(* IEC 61131-3 sources: T4Exjobb/Sigma/Stations/MachineControl/MachineControl/Network, 1 file *)

(* ---- ConfigObjects.st ---- *)
FUNCTION GLOBAL TAB TASK_CONF
_K_TASK, _K_REAL,
_K_END_VAR,

_K_TASK, _K_CYCLIC,
_K_END_VAR,

_K_TASK, _K_BACKGROUND,
_K_END_VAR,

_K_END_CONF
END_FUNCTION

FUNCTION GLOBAL TAB IPR_CONF
_K_IPR
	0$UINT,
_K_END_VAR,
_K_END_CONF
END_FUNCTION

FUNCTION GLOBAL TAB CONFIG_TABLES
00034$UINT,
0$UINT, 0, 11, "_ALARMX0PARA",
0$UINT, 0, 19, "_ALARMXBUFFER",
0$UINT, 1, 3, "_CHECKONLINESTATUS",
0$UINT, 1, 0, "_CHECKSUM",
0$UINT, 1, 1, "_MULTITASK",
0$UINT, 1, 0, "_SIG_LSL_CMULTIMASTERSTATE",
0$UINT, 0, 0, "_STDLIB",
0$UINT, 2, 0, "_SYNCTIMEPLC",
0$UINT, 0, 7, "_SYSDATETIME",
0$UINT, 0, 0, "_SYSDATETIME2",
0$UINT, 1, 1, "_TASKOBJECTCONTROL",
0$UINT, 1, 17, "_TCPIP_CLIENT",
0$UINT, 1, 36, "_TCPIP_SERVER",
0$UINT, 1, 20, "ASCII_BIN",
0$UINT, 0, 4, "CRITICALSECTION",
0$UINT, 1, 0, "DATAMANAGER",
0$UINT, 1, 0, "DATAMANAGERFIFO",
0$UINT, 1, 0, "DATAMANAGERPRIORITY",
0$UINT, 1, 2, "GETOSVERSION",
0$UINT, 0, 2, "GETTASKHANDLE",
0$UINT, 1, 22, "MERKEREX",
0$UINT, 1, 68, "PLC_INFO",
0$UINT, 1, 3, "RAM",
0$UINT, 1, 1, "RAMRINGBUFFER",
0$UINT, 0, 0, "READER",
0$UINT, 0, 23, "SIGCLIB",
0$UINT, 1, 10, "STRING",
0$UINT, 1, 82, "STRINGINTERNAL",
0$UINT, 0, 1, "SYSTEM",
0$UINT, 1, 14, "TCPCOMMUNICATION",
0$UINT, 1, 0, "TCPCOMMUNICATIONLOGFILTER",
0$UINT, 0, 0, "TCPV2",
0$UINT, 1, 1, "USERALARMGENERATOR",
0$UINT, 1, 3, "VIRTUALBASEINIT",
ONE_CFG$UINT, 0, 0, "ONE_Main",
ONE_CFG$UINT, 1, 0, "ONE_STDAlarm",
ONE_CFG$UINT, 1, 0, "ONE_STDCommunicationToHMI",
ONE_CFG$UINT, 1, 0, "ONE_STDPLCInfoPLC",
ONE_CFG$UINT, 2, 0, "ONE_STDTimeSync",
TASK_CFG$UINT, 0, 0, "TASK_CONF",
IPR_CFG$UINT, 0, 0, "IPR_CONF",
PRJ_CFG$UINT, 0, 0, "MachineControl",
END_FUNCTION

FUNCTION GLOBAL TAB CH_REDIRECT_EMB_TAB
0000$UINT,
00015$UINT,
"_TCPIP_CLIENT;SemaName01", "\StrSemaName01.Data",
"_TCPIP_CLIENT;SemaName02", "\StrSemaName02.Data",
"_TCPIP_CLIENT;TaskName", "\StrTaskName.Data",
"_TCPIP_SERVER;SemaName01", "\StrSemaName01.Data",
"_TCPIP_SERVER;SemaName02", "\StrSemaName02.Data",
"_TCPIP_SERVER;TaskName", "\StrTaskName.Data",
"PLC_Info;ApplicationName", "\AppliName.Data",
"PLC_Info;CPUBoardName", "\CPUBoard.Data",
"PLC_Info;CPU_Name", "\String1.Data",
"PLC_Info;SerNum", "\String0.Data",
"PLC_Info;SysInfoString", "\SysInfo.Data",
"Reader;SemaName01", "\StrSemaName01.Data",
"Reader;SemaName02", "\StrSemaName02.Data",
"Reader;TaskName", "\StrTaskName.Data",
"TCPCommunication;TaskName", "\ThreadName.Data",
END_FUNCTION
